FUNCTION_BLOCK DEMUX (* Composite Function Block Type *)
  (* Standard: 61499-2 *)
  (* Version 0.0, 10/11/2026, macie, nxtControl GmBH, template *)
  PACKAGE Main;
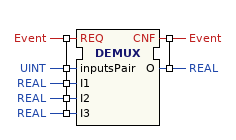
  EVENT_INPUT
    REQ WITH inputsPair, I1, I2, I3; (* Normal Execution Request *)
  END_EVENT
  EVENT_OUTPUT
    CNF WITH O; (* Execution Confirmation *)
  END_EVENT
  VAR_INPUT
    inputsPair : UINT;
    I1 : REAL; (* Input event qualifier *)
    I2 : REAL;
    I3 : REAL;
  END_VAR
  VAR_OUTPUT
    O : REAL; (* Output event qualifier *)
  END_VAR
END_FUNCTION_BLOCK
